Fanuc KAREL source: kc00060.KL

-- PROVISIONAL review KL for V1013-1; original PC SHA256 60c8fe4e7f07f425fd340d41753292bd791505d4afd96928212b1850bddfd139
-- Incomplete behavior may be omitted. Consult companion uncertainty JSON. Do not deploy.
PROGRAM KC00060
%NOLOCKGROUP
BEGIN
  -- UNRESOLVED_PC offsets 5-43; opcodes 27,27,9D,22,1C,22,22,2A,AA,23
  -- UNRESOLVED_PC offsets 48-52; opcodes 7F
END KC00060
